Yaskawa INFORM job: SLINJE1.JBI

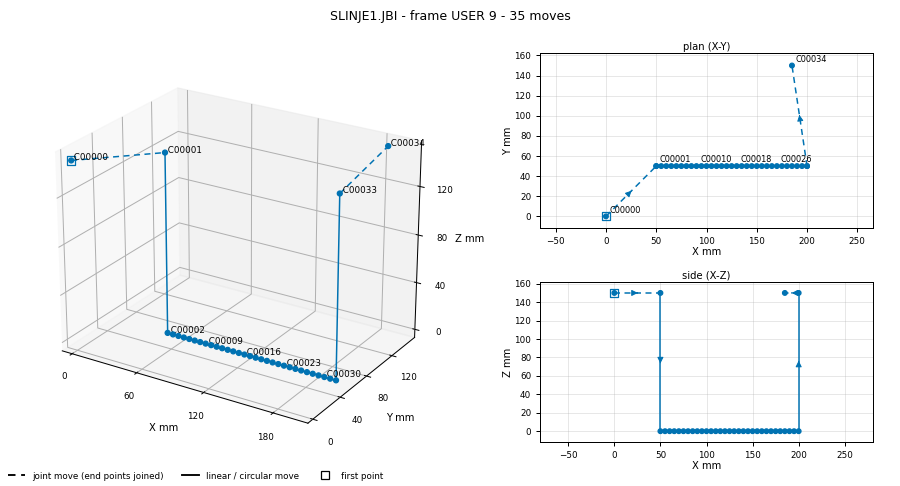
[picture p0: tool path of SLINJE1.JBI in frame USER 9, 35 of 35 moves have a stored position in this frame; points joined in program order, loops and branches not executed]
/JOB
//NAME SLINJE1
//POS
///NPOS 35,0,0,0,0,0
///USER 9
///TOOL 1
///POSTYPE USER
///RECTAN
///RCONF 1,0,0,0,0,0,0,0,0,0,0,0,0,0,0,0,0,0,0,0,0,0,0,0
C00000=0.000,0.000,150.000,0.0000,0.0000,180.0000
C00001=50.000,50.000,150.000,0.0000,0.0000,180.0000
C00002=50.000,50.000,0.000,0.0000,0.0000,180.0000
C00003=55.000,50.000,0.000,0.0000,0.0000,180.0000
C00004=60.000,50.000,0.000,0.0000,0.0000,180.0000
C00005=65.000,50.000,0.000,0.0000,0.0000,180.0000
C00006=70.000,50.000,0.000,0.0000,0.0000,180.0000
C00007=75.000,50.000,0.000,0.0000,0.0000,180.0000
C00008=80.000,50.000,0.000,0.0000,0.0000,180.0000
C00009=85.000,50.000,0.000,0.0000,0.0000,180.0000
C00010=90.000,50.000,0.000,0.0000,0.0000,180.0000
C00011=95.000,50.000,0.000,0.0000,0.0000,180.0000
C00012=100.000,50.000,0.000,0.0000,0.0000,180.0000
C00013=105.000,50.000,0.000,0.0000,0.0000,180.0000
C00014=110.000,50.000,0.000,0.0000,0.0000,180.0000
C00015=115.000,50.000,0.000,0.0000,0.0000,180.0000
C00016=120.000,50.000,0.000,0.0000,0.0000,180.0000
C00017=125.000,50.000,0.000,0.0000,0.0000,180.0000
C00018=130.000,50.000,0.000,0.0000,0.0000,180.0000
C00019=135.000,50.000,0.000,0.0000,0.0000,180.0000
C00020=140.000,50.000,0.000,0.0000,0.0000,180.0000
C00021=145.000,50.000,0.000,0.0000,0.0000,180.0000
C00022=150.000,50.000,0.000,0.0000,0.0000,180.0000
C00023=155.000,50.000,0.000,0.0000,0.0000,180.0000
C00024=160.000,50.000,0.000,0.0000,0.0000,180.0000
C00025=165.000,50.000,0.000,0.0000,0.0000,180.0000
C00026=170.000,50.000,0.000,0.0000,0.0000,180.0000
C00027=175.000,50.000,0.000,0.0000,0.0000,180.0000
C00028=180.000,50.000,0.000,0.0000,0.0000,180.0000
C00029=185.000,50.000,0.000,0.0000,0.0000,180.0000
C00030=190.000,50.000,0.000,0.0000,0.0000,180.0000
C00031=195.000,50.000,0.000,0.0000,0.0000,180.0000
C00032=200.000,50.000,0.000,0.0000,0.0000,180.0000
C00033=200.000,50.000,150.000,0.0000,0.0000,180.0000
C00034=185.000,150.000,150.000,0.0000,0.0000,180.0000
//INST
///DATE 2026/10/20 11:28
///ATTR SC,RW,RJ
////FRAME USER 9
///GROUP1 RB1
NOP
MOVJ C00000 VJ=0.78
MOVJ C00001 VJ=0.78
MOVL C00002 V=11.0 ACC=20 DEC=20
MACRO1 MJ#(0) ARGF205
ARCON
MOVL C00003 V=8.0 ACC=20 DEC=20
MOVL C00004 V=8.0 ACC=20 DEC=20
MOVL C00005 V=8.0 ACC=20 DEC=20
MOVL C00006 V=8.0 ACC=20 DEC=20
MOVL C00007 V=8.0 ACC=20 DEC=20
MOVL C00008 V=8.0 ACC=20 DEC=20
MOVL C00009 V=8.0 ACC=20 DEC=20
MOVL C00010 V=8.0 ACC=20 DEC=20
MOVL C00011 V=8.0 ACC=20 DEC=20
MOVL C00012 V=8.0 ACC=20 DEC=20
MOVL C00013 V=8.0 ACC=20 DEC=20
MOVL C00014 V=8.0 ACC=20 DEC=20
MOVL C00015 V=8.0 ACC=20 DEC=20
MOVL C00016 V=8.0 ACC=20 DEC=20
MOVL C00017 V=8.0 ACC=20 DEC=20
MOVL C00018 V=8.0 ACC=20 DEC=20
MOVL C00019 V=8.0 ACC=20 DEC=20
MOVL C00020 V=8.0 ACC=20 DEC=20
MOVL C00021 V=8.0 ACC=20 DEC=20
MOVL C00022 V=8.0 ACC=20 DEC=20
MOVL C00023 V=8.0 ACC=20 DEC=20
MOVL C00024 V=8.0 ACC=20 DEC=20
MOVL C00025 V=8.0 ACC=20 DEC=20
MOVL C00026 V=8.0 ACC=20 DEC=20
MOVL C00027 V=8.0 ACC=20 DEC=20
MOVL C00028 V=8.0 ACC=20 DEC=20
MOVL C00029 V=8.0 ACC=20 DEC=20
MOVL C00030 V=8.0 ACC=20 DEC=20
MOVL C00031 V=8.0 ACC=20 DEC=20
MOVL C00032 V=8.0 ACC=20 DEC=20
ARCOF
MOVL C00033 V=11.0 ACC=20 DEC=20
MOVJ C00034 VJ=0.78
END
